// TIA Portal V21 export
FUNCTION_BLOCK "LadLogic"   // FB10, LAD
TITLE = Ladder logic
{ S7_Optimized_Access := 'TRUE' }
// Bit logic in ladder: contacts, coils, an edge and a jump.
   VAR_INPUT
      start : Bool;
      stop : Bool;
      door : Bool;
   END_VAR
   VAR_OUTPUT
      motor : Bool;
      lamp : Bool;
      fault : Bool;
   END_VAR
   VAR
      latched : Bool;
      edgeMemory : Bool;
   END_VAR
   VAR_TEMP   // added for the SCL form of the ladder/FBD networks
      _w1 : Bool;
   END_VAR
BEGIN

REGION Network 1: Start and stop
   // Contacts in series and in parallel drive the motor.
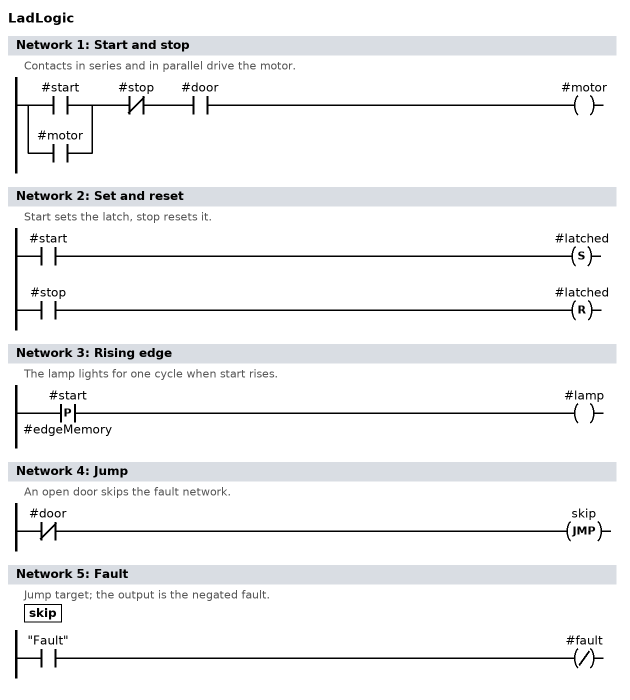
   #motor := (#start OR #motor) AND NOT #stop AND #door;
END_REGION

REGION Network 2: Set and reset
   // Start sets the latch, stop resets it.
   RUNG wire#powerrail
      Contact( #start )
      S_Coil( #latched )
   END_RUNG
   RUNG wire#powerrail
      Contact( #stop )
      R_Coil( #latched )
   END_RUNG
   // the same network as SCL:
   IF #start THEN #latched := TRUE; END_IF;
   IF #stop THEN #latched := FALSE; END_IF;
END_REGION

REGION Network 3: Rising edge
   // The lamp lights for one cycle when start rises.
   RUNG wire#powerrail
      P_Contact(operand := #start, bit := #edgeMemory)
      Coil( #lamp )
   END_RUNG
   // the same network as SCL:
   #_w1 := #start AND NOT #edgeMemory;   // rising edge of #start
   #edgeMemory := #start;
   #lamp := #_w1;
END_REGION

REGION Network 4: Jump
   // An open door skips the fault network.
   RUNG wire#powerrail
      I_Contact( #door )
      JumpCoil( skip )
   END_RUNG
   // the same network as SCL:
   IF NOT #door THEN GOTO skip; END_IF;
END_REGION

REGION Network 5: Fault
   // Jump target; the output is the negated fault.
   Label( skip )
   RUNG wire#powerrail
      Contact( "Fault" )
      I_Coil( #fault )
   END_RUNG
   // the same network as SCL:
   skip:
   #fault := NOT "Fault";
END_REGION
END_FUNCTION_BLOCK
